FUNCTION_BLOCK Motor_Generico_HMI (* Service Interface Function Block Type *)
  (* Standard: 61499-2 *)
  (* Version 1.8, 21/10/2026, Hidryco, Hidryco, IHM do Motor_Generico 1.8: STS_FALHA = falha ativa *)
  PACKAGE Hidryco.HidrycoLib;
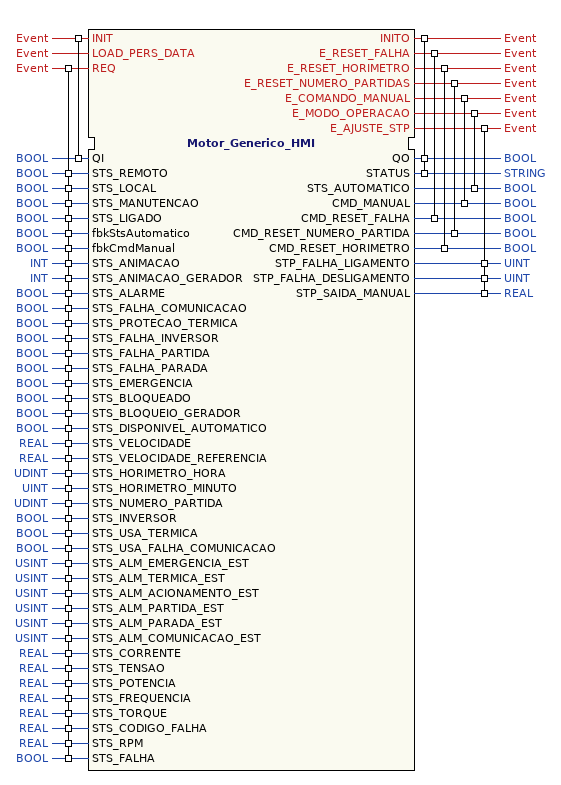
  EVENT_INPUT
    INIT WITH QI;
    LOAD_PERS_DATA; (* Reenvia os parametros persistentes *)
    REQ WITH STS_REMOTO, STS_LOCAL, STS_MANUTENCAO, STS_LIGADO, fbkStsAutomatico, fbkCmdManual, STS_ANIMACAO, STS_ANIMACAO_GERADOR, STS_ALARME, STS_FALHA_COMUNICACAO, STS_PROTECAO_TERMICA, STS_FALHA_INVERSOR, STS_FALHA_PARTIDA, STS_FALHA_PARADA, STS_EMERGENCIA, STS_BLOQUEADO, STS_BLOQUEIO_GERADOR, STS_DISPONIVEL_AUTOMATICO, STS_VELOCIDADE, STS_VELOCIDADE_REFERENCIA, STS_HORIMETRO_HORA, STS_HORIMETRO_MINUTO, STS_NUMERO_PARTIDA, STS_INVERSOR, STS_USA_TERMICA, STS_USA_FALHA_COMUNICACAO, STS_ALM_EMERGENCIA_EST, STS_ALM_TERMICA_EST, STS_ALM_ACIONAMENTO_EST, STS_ALM_PARTIDA_EST, STS_ALM_PARADA_EST, STS_ALM_COMUNICACAO_EST, STS_CORRENTE, STS_TENSAO, STS_POTENCIA, STS_FREQUENCIA, STS_TORQUE, STS_CODIGO_FALHA, STS_RPM, STS_FALHA; (* Atualizacao de status *)
  END_EVENT
  EVENT_OUTPUT
    INITO WITH QO, STATUS;
    E_RESET_FALHA WITH CMD_RESET_FALHA;
    E_RESET_HORIMETRO WITH CMD_RESET_HORIMETRO;
    E_RESET_NUMERO_PARTIDAS WITH CMD_RESET_NUMERO_PARTIDA;
    E_COMANDO_MANUAL WITH CMD_MANUAL;
    E_MODO_OPERACAO WITH STS_AUTOMATICO;
    E_AJUSTE_STP WITH STP_FALHA_LIGAMENTO, STP_FALHA_DESLIGAMENTO, STP_SAIDA_MANUAL;
  END_EVENT
  VAR_INPUT
    QI : BOOL;
    STS_REMOTO : BOOL; (* Chave em remoto *)
    STS_LOCAL : BOOL; (* Chave em local *)
    STS_MANUTENCAO : BOOL; (* Chave nem local nem remoto *)
    STS_LIGADO : BOOL; (* Motor ligado *)
    fbkStsAutomatico : BOOL; (* Modo automatico (retorno para a IHM) *)
    fbkCmdManual : BOOL; (* Comando manual em vigor (retorno para a IHM) *)
    STS_ANIMACAO : INT; (* 0 desligado, 1 ligado, 2 falha, 3 manutencao *)
    STS_ANIMACAO_GERADOR : INT; (* 0 nao conectado, 1 conectado, 2 selecionado, 3 selecionado e gerador ligado *)
    STS_ALARME : BOOL; (* Alarme geral *)
    STS_FALHA_COMUNICACAO : BOOL; (* Falha de comunicacao com a remota *)
    STS_PROTECAO_TERMICA : BOOL; (* Falha termica (memorizada) *)
    STS_FALHA_INVERSOR : BOOL; (* Falha do inversor/acionamento (memorizada) *)
    STS_FALHA_PARTIDA : BOOL; (* Nao confirmou partida (memorizada) *)
    STS_FALHA_PARADA : BOOL; (* Nao confirmou parada (memorizada) *)
    STS_EMERGENCIA : BOOL; (* Emergencia (memorizada) *)
    STS_BLOQUEADO : BOOL; (* Intertravamento ativo *)
    STS_BLOQUEIO_GERADOR : BOOL; (* Bloqueado pelo gerador *)
    STS_DISPONIVEL_AUTOMATICO : BOOL; (* Disponivel para o automatico *)
    STS_VELOCIDADE : REAL; (* Velocidade (%): com inversor 0 % no LSP e 100 % no HSP; sem inversor 0 ou 100 *)
    STS_VELOCIDADE_REFERENCIA : REAL; (* Referencia de velocidade (Hz) *)
    STS_HORIMETRO_HORA : UDINT; (* Horimetro (h) *)
    STS_HORIMETRO_MINUTO : UINT; (* Horimetro (min) *)
    STS_NUMERO_PARTIDA : UDINT; (* Numero de partidas *)
    STS_INVERSOR : BOOL; (* Motor com inversor *)
    STS_USA_TERMICA : BOOL; (* Configuracao: termica supervisionada (IHM mostra a linha da termica) *)
    STS_USA_FALHA_COMUNICACAO : BOOL; (* Configuracao: falha de comunicacao supervisionada *)
    STS_ALM_EMERGENCIA_EST : USINT; (* Estado do ALARM_BIT (0 normal, 1 ativo reconhecido, 2 ativo nao reconhecido, 3 saiu nao reconhecido, 4 ativo e saiu nao reconhecido) *)
    STS_ALM_TERMICA_EST : USINT; (* Estado do ALARM_BIT (0 normal, 1 ativo reconhecido, 2 ativo nao reconhecido, 3 saiu nao reconhecido, 4 ativo e saiu nao reconhecido) *)
    STS_ALM_ACIONAMENTO_EST : USINT; (* Estado do ALARM_BIT (0 normal, 1 ativo reconhecido, 2 ativo nao reconhecido, 3 saiu nao reconhecido, 4 ativo e saiu nao reconhecido) *)
    STS_ALM_PARTIDA_EST : USINT; (* Estado do ALARM_BIT (0 normal, 1 ativo reconhecido, 2 ativo nao reconhecido, 3 saiu nao reconhecido, 4 ativo e saiu nao reconhecido) *)
    STS_ALM_PARADA_EST : USINT; (* Estado do ALARM_BIT (0 normal, 1 ativo reconhecido, 2 ativo nao reconhecido, 3 saiu nao reconhecido, 4 ativo e saiu nao reconhecido) *)
    STS_ALM_COMUNICACAO_EST : USINT; (* Estado do ALARM_BIT (0 normal, 1 ativo reconhecido, 2 ativo nao reconhecido, 3 saiu nao reconhecido, 4 ativo e saiu nao reconhecido) *)
    STS_CORRENTE : REAL; (* Corrente (A) *)
    STS_TENSAO : REAL; (* Tensao (V) *)
    STS_POTENCIA : REAL; (* Potencia (kW) *)
    STS_FREQUENCIA : REAL; (* Frequencia (Hz) *)
    STS_TORQUE : REAL; (* Torque (%) *)
    STS_CODIGO_FALHA : REAL; (* Codigo de falha do inversor *)
    STS_RPM : REAL; (* Rotacao (rpm) *)
    STS_FALHA : BOOL; (* Falha ativa: motor em falha agora (emergencia, termica, acionamento ou comunicacao), sem memoria *)
  END_VAR
  VAR_OUTPUT
    QO : BOOL; (* Event Output Qualifier *)
    STATUS : STRING; (* Service Status *)
    STS_AUTOMATICO : BOOL; (* 0 = manual, 1 = automatico (persistente) *)
    CMD_MANUAL : BOOL; (* 0 = desligar, 1 = ligar (nao persistente) *)
    CMD_RESET_FALHA : BOOL; (* Reset de falhas *)
    CMD_RESET_NUMERO_PARTIDA : BOOL; (* Zera numero de partidas *)
    CMD_RESET_HORIMETRO : BOOL; (* Zera horimetro *)
    STP_FALHA_LIGAMENTO : UINT; (* Tempo maximo para confirmar partida (s). 0 = desabilitado *)
    STP_FALHA_DESLIGAMENTO : UINT; (* Tempo maximo para confirmar parada (s). 0 = desabilitado *)
    STP_SAIDA_MANUAL : REAL; (* Velocidade em manual (Hz) *)
  END_VAR
  SERVICE /
    SEQUENCE 
    END_SEQUENCE
  END_SERVICE
END_FUNCTION_BLOCK
